FUNCTION_BLOCK Desinfeccao_UV (* Desinfeccao UV e limitacao da vazao de lancamento (700) - HidrycoLib *)
  (* Standard: 61499-2 *)
  (* Version 1.3, 21/10/2026, Hidryco, Hidryco, 1.3: REQ_GERADOR (geradorHabilitaUV01/02, stsGerador; Subestacao HAB_UV_700_01/02 e stsPlantaNoGerador) repassado ao UV para o raio dos canais. 1.2: pidCtl Pid com CycleTime 1000 ms (sem ele o calculo ciclico do pidSC ficava sem periodo). 1.1: ajustes do PID no sub-CAT PID_VC_700_01 (padrao Desinfeccao do legado; desejado = vazao maxima); reset cmdResetFalhas / E_RESET_FALHAS_PROCESSO; AIT_700_01/03/04. 1.0: desinfeccao (700). Sub-CATs: VC_700_01 (Valvula_Coester modulante), UV (UV_Trojan), FT_700_01 (Parshall 4-20 mA, m3/h), AIT_700_001 turbidez, AIT_700_003 pH, AIT_700_004 OD (SC4500 por comunicacao). PID continuo (pidCtl, Direction TRUE: vazao acima do setpoint fecha a valvula) limita a vazao de lancamento (padrao 1242 m3/h = 345 L/s). Campo por symlink ${PATH}: djPCEDesligado, djPCMDesligado, djUV01, djUV02, djVC01, djMO01 (remota %I0.0-0.5), stsRemotaComOk (COM_OK do IO_DI32 da remota). *)
  PACKAGE Hidryco.HidrycoLib;
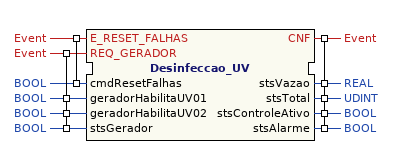
  EVENT_INPUT
    E_RESET_FALHAS WITH cmdResetFalhas; (* Reset pelo processo (desinfeccao, valvula, UV e sensores) com cmdResetFalhas = TRUE *)
    REQ_GERADOR WITH geradorHabilitaUV01, geradorHabilitaUV02, stsGerador; (* Planta no gerador e liberacao do UV (Subestacao) *)
  END_EVENT
  EVENT_OUTPUT
    CNF WITH stsVazao, stsTotal, stsControleAtivo, stsAlarme; (* Status *)
  END_EVENT
  VAR_INPUT
    cmdResetFalhas : BOOL; (* TRUE = reset (com o evento E_RESET_FALHAS) *)
    geradorHabilitaUV01 : BOOL; (* 700-UV-01 liberado para operar com a planta nos geradores *)
    geradorHabilitaUV02 : BOOL; (* 700-UV-02 liberado para operar com a planta nos geradores *)
    stsGerador : BOOL; (* TRUE = planta alimentada pelos geradores *)
  END_VAR
  VAR_OUTPUT
    stsVazao : REAL; (* Vazao do efluente final (m3/h) *)
    stsTotal : UDINT; (* Volume totalizado (m3) *)
    stsControleAtivo : BOOL; (* PID controlando a 700-VC-01 *)
    stsAlarme : BOOL; (* Algum alarme da desinfeccao *)
  END_VAR
  FBS
    IThis : Desinfeccao_UV_HMI(QI := TRUE);
    plcStart1 : plcStart(Prio := 10);
    Logica : basicDesinfeccao;
    Tick : E_CYCLE(DT := T#1s);
    Pid : pidCtl(CycleTime := 1000, Direction := TRUE, Bump := FALSE, ProhibitOutInc := FALSE, ProhibitOutDec := FALSE);
    PersTotal : PERSISTENCE_20652AC5DB8BA8AD5(QI := TRUE); {SET_ATTRIBUTE(Configuration.GenericFBType.InterfaceParams, Runtime.Standard#I:=3;input${I$}:UINT,UINT,UDINT)}
    Disjuntores : SYMLINKMULTIVARDST_5495E501E675F500(QI := TRUE, NAME1 := '$${PATH}djPCEDesligado', NAME2 := '$${PATH}djPCMDesligado', NAME3 := '$${PATH}djUV01', NAME4 := '$${PATH}djUV02', NAME5 := '$${PATH}djVC01', NAME6 := '$${PATH}djMO01'); {SET_ATTRIBUTE(Configuration.GenericFBType.InterfaceParams, Runtime.System#I:=6;VALUE${I$}:BOOL,BOOL,BOOL,BOOL,BOOL,BOOL)}
    Remota : SYMLINKMULTIVARDST_1559B0FF8170C9BA0(QI := TRUE, NAME1 := '$${PATH}stsRemotaComOk'); {SET_ATTRIBUTE(Configuration.GenericFBType.InterfaceParams, Runtime.System#I:=1;VALUE${I$}:BOOL)}
    FT_700_01 : Sensor_Generico(pin_CC8EEC06FF0C4430 := 'm3/h', pin_6D3A2524C5D0F0D1 := 0);
    AIT_700_01 : Sensor_Generico(pin_D46B37D45FD5AF5D := TRUE, pin_0ECE7B3867B02E0B := TRUE, pin_CC8EEC06FF0C4430 := 'NTU', pin_6D3A2524C5D0F0D1 := 1);
    AIT_700_03 : Sensor_Generico(pin_D46B37D45FD5AF5D := TRUE, pin_0ECE7B3867B02E0B := TRUE, pin_CC8EEC06FF0C4430 := '', pin_6D3A2524C5D0F0D1 := 2);
    AIT_700_04 : Sensor_Generico(pin_D46B37D45FD5AF5D := TRUE, pin_CC8EEC06FF0C4430 := 'mV', pin_6D3A2524C5D0F0D1 := 0); (* ORP (mV) do SC4500 de pH (conexao supervisionada pelo AIT_700_03: o connStatusInt so tem um destino) *)
    VC_700_01 : Atuador_Coester(pin_C65F121E4D57852C := TRUE);
    UV : UV_Trojan;
    AlarmeVazaoAlta : ALARM_BIT(TYPE := 1, ACKTYPE_1 := 2, ACTIVE := TRUE); {SET_ATTRIBUTE(HMI.AlarmText, Vazão de lançamento acima do limite)}
    AlarmeVariacao : ALARM_BIT(TYPE := 1, ACKTYPE_1 := 2, ACTIVE := TRUE); {SET_ATTRIBUTE(HMI.AlarmText, Variação brusca da vazão de lançamento)} {SET_ATTRIBUTE(HMI.AlarmClass, Warning)}
    AlarmeDisjuntor : ALARM_BIT(TYPE := 1, ACKTYPE_1 := 2, ACTIVE := TRUE); {SET_ATTRIBUTE(HMI.AlarmText, Disjuntor da desinfecção desligado)} {SET_ATTRIBUTE(HMI.AlarmClass, Warning)}
    AlarmeRemota : ALARM_BIT(TYPE := 1, ACKTYPE_1 := 2, ACTIVE := TRUE); {SET_ATTRIBUTE(HMI.AlarmText, Remota da desinfecção sem comunicação)} {SET_ATTRIBUTE(HMI.AlarmClass, Warning)}
    PID_VC_700_01 : Controle_PID;
  END_FBS
  EVENT_CONNECTIONS
    plcStart1.FIRST_INIT TO IThis.B18F9527B03F6368;
    plcStart1.REDO_INIT TO IThis.B18F9527B03F6368;
    IThis.8DA18C8B88D861AA TO Disjuntores.INIT;
    Disjuntores.INITO TO Remota.INIT;
    Remota.INITO TO Logica.9E12B42E11EB9FB7;
    Remota.INITO TO IThis.B29E261CF0325DC9;
    Logica.39B67DFC9697D1D0 TO Tick.START;
    Logica.39B67DFC9697D1D0 TO PersTotal.INIT;
    PersTotal.INITO TO PersTotal.READ;
    PersTotal.READCNF TO Logica.2E96492E37281113;
    Logica.BC4C937414AD6E45 TO PersTotal.WRITE;
    Logica.39B67DFC9697D1D0 TO AlarmeVazaoAlta.INIT;
    AlarmeVazaoAlta.INITO TO AlarmeVazaoAlta.REQ_INITDATA;
    AlarmeVazaoAlta.CNF_INITDATA TO AlarmeVazaoAlta.ACTIVATE;
    AlarmeVariacao.INITO TO AlarmeVariacao.REQ_INITDATA;
    AlarmeVariacao.CNF_INITDATA TO AlarmeVariacao.ACTIVATE;
    AlarmeVazaoAlta.INITO TO AlarmeVariacao.INIT;
    AlarmeDisjuntor.INITO TO AlarmeDisjuntor.REQ_INITDATA;
    AlarmeDisjuntor.CNF_INITDATA TO AlarmeDisjuntor.ACTIVATE;
    AlarmeVariacao.INITO TO AlarmeDisjuntor.INIT;
    AlarmeRemota.INITO TO AlarmeRemota.REQ_INITDATA;
    AlarmeRemota.CNF_INITDATA TO AlarmeRemota.ACTIVATE;
    AlarmeDisjuntor.INITO TO AlarmeRemota.INIT;
    AlarmeRemota.INITO TO plcStart1.ACK_FIRST;
    Tick.EO TO Logica.A43A58424E0F5DF5;
    Disjuntores.CNF TO Logica.22B807AE7A8B903D;
    Remota.CNF TO Logica.2AE8EBA1815E0012;
    FT_700_01.28A380156DB271B8 TO Logica.6559A273E8431D42;
    VC_700_01.CF6616D3CB5312F6 TO Logica.4F5B69463931E86B;
    UV.41148E14CCAE49D5 TO Logica.1495D2B4E524DEC3;
    Logica.6010724B5A00E1A3 TO VC_700_01.6AE7937B5439A162;
    FT_700_01.28A380156DB271B8 TO Pid.REQ;
    Logica.38355A458523F08C TO Pid.REQ;
    Pid.CNF TO Logica.1DD56BE62400BF1C;
    Pid.C_CNF TO Logica.1DD56BE62400BF1C;
    IThis.341E4C9D143B2914 TO Logica.69B239DBC6B5BF03;
    IThis.673C9CACFA30E81B TO Logica.F980CDC9B2AFA9D8;
    IThis.A7123D0B6BA18805 TO Logica.B454118112B7B3A8;
    Logica.04CB25776C0D242A TO IThis.1B47BC94CEE432D9;
    Logica.04CB25776C0D242A TO AlarmeVazaoAlta.REQ;
    AlarmeVazaoAlta.IND_1 TO IThis.1B47BC94CEE432D9;
    IThis.673C9CACFA30E81B TO AlarmeVazaoAlta.ACK_C1;
    Logica.04CB25776C0D242A TO AlarmeVariacao.REQ;
    AlarmeVariacao.IND_1 TO IThis.1B47BC94CEE432D9;
    IThis.673C9CACFA30E81B TO AlarmeVariacao.ACK_C1;
    Logica.04CB25776C0D242A TO AlarmeDisjuntor.REQ;
    AlarmeDisjuntor.IND_1 TO IThis.1B47BC94CEE432D9;
    IThis.673C9CACFA30E81B TO AlarmeDisjuntor.ACK_C1;
    Logica.04CB25776C0D242A TO AlarmeRemota.REQ;
    AlarmeRemota.IND_1 TO IThis.1B47BC94CEE432D9;
    IThis.673C9CACFA30E81B TO AlarmeRemota.ACK_C1;
    E_RESET_FALHAS TO Logica.DA13244B5D56E79F;
    E_RESET_FALHAS TO FT_700_01.D21DAA5004F58516;
    E_RESET_FALHAS TO AIT_700_01.D21DAA5004F58516;
    E_RESET_FALHAS TO AIT_700_03.D21DAA5004F58516;
    E_RESET_FALHAS TO AIT_700_04.D21DAA5004F58516;
    E_RESET_FALHAS TO VC_700_01.D903CD18EBE204D1;
    Logica.6AA932C3761CE99C TO CNF;
    PID_VC_700_01.75EB05A15DC6DC61 TO Pid.REQ_PARA;
    PID_VC_700_01.75EB05A15DC6DC61 TO Pid.REQ_SP;
    PID_VC_700_01.75EB05A15DC6DC61 TO Logica.69B239DBC6B5BF03;
    Remota.INITO TO PID_VC_700_01.117942CC3F34C94C;
    Logica.04CB25776C0D242A TO PID_VC_700_01.7BD84B0FC1882775;
    REQ_GERADOR TO UV.6FAFCDDE653CB65D;
  END_CONNECTIONS
  DATA_CONNECTIONS
    PersTotal.output3 TO Logica.E77A551E7F1625D6;
    Logica.BB35FC69145014F5 TO PersTotal.input3;
    Disjuntores.VALUE1 TO Logica.CF45361D95BFAA25;
    Disjuntores.VALUE2 TO Logica.347EEF72575B0DAD;
    Disjuntores.VALUE3 TO Logica.159FAE7A20FE4F43;
    Disjuntores.VALUE4 TO Logica.7868F97BB44D7BB6;
    Disjuntores.VALUE5 TO Logica.92824DDB3BCC4699;
    Disjuntores.VALUE6 TO Logica.50FED92E4734ACF3;
    Remota.VALUE1 TO Logica.D0484A6EFE322016;
    FT_700_01.D7422D307E6AF52D TO Logica.F569AB39D886D3C5;
    FT_700_01.726640D1704B3F86 TO Logica.8F6D70C85B5729EE;
    VC_700_01.904DD3246D8E0F2F TO Logica.C5936F826382DFB8;
    VC_700_01.259F220E31BE1DFA TO Logica.7315FEF776808725;
    VC_700_01.5B46E3B5D12031DA TO Logica.023A1B52E4E2056D;
    VC_700_01.378CDAA06C4824E3 TO Logica.DBD5C62FC984909D;
    UV.8A986F32247F8461 TO Logica.DB1DCC8BAF4C9029;
    UV.EDFBC67855FC1BF4 TO Logica.1AFFBF765DAF6E05;
    UV.53F24ADA26C29448 TO Logica.6927441A48A28A44;
    UV.E73DB33437F0D160 TO Logica.FA4C9F16C9AD1E00;
    UV.B5E6F2B1B4A7F74D TO Logica.E17D46372D8AC1CC;
    UV.2373201554B21091 TO Logica.CA02F082C523342B;
    Logica.635B91EC32B193D8 TO VC_700_01.B08C4ED4004BD1E2;
    FT_700_01.D7422D307E6AF52D TO Pid.Pv;
    Logica.B925699CCA1010B0 TO Pid.Mode;
    Logica.E0C52E4AA1CB94A3 TO Pid.PresetValue;
    Pid.Out TO Logica.AA3C6B9770CFA1D6;
    IThis.975D7F4B71294A99 TO Logica.A62BE056EBF6633F;
    IThis.48B1DA7F68ECA0A8 TO Logica.0CA93D1DC0F0D80A;
    IThis.BF0DC1C37334FADC TO Logica.EAB397A6710197DE;
    IThis.3223A03025B9D306 TO Logica.14F8441489A49AD8;
    IThis.133D4C207A85139E TO Logica.EDA9F4A4D8516735;
    Logica.8B489663C97AF746 TO IThis.64C5B4D669700647;
    Logica.2CB6FFAA3F88FD37 TO IThis.9BBBF4F79C014F9D;
    Logica.1AC4273BD48629B4 TO IThis.ED2A3A2AD9D2CEAB;
    Logica.7C47B967196CD681 TO IThis.8CFA6BB1EE69DBDA;
    Logica.F5E44B9CD467E225 TO IThis.9D544CFE60C51E40;
    Logica.E0E853656DE9663A TO IThis.00083F484189930B;
    Logica.5B994E1E72A57859 TO IThis.5A630CE8F223E31A;
    Logica.9D46B9FE82DC9AB1 TO IThis.3724F9189B78EC4D;
    Logica.06E435E0579C0A31 TO IThis.4C496D880FB42A44;
    Logica.03E13841379C7979 TO IThis.DE11125D4105DF0E;
    Logica.9EE277DF1A6EE639 TO IThis.909A978770157DD8;
    Logica.DD39785BA0B3D6D1 TO IThis.D8676A9461C485D9;
    Logica.DC6A854DD28F4447 TO IThis.8155290424886535;
    Logica.CFF2FF9B070BCB84 TO IThis.E0FD426C54E10B50;
    Logica.A1948102A71BA04F TO IThis.B5278628A6F4EB0E;
    Logica.49CC92A2C50C5502 TO IThis.3146A9607323897C;
    Logica.029A5972D76D7D9D TO IThis.207239DB8C69408E;
    Logica.7C31ABB79E620CA1 TO IThis.0DCEC12DB41BD8A9;
    Logica.4979C9EBFE656646 TO IThis.F89132E9AC0FBE71;
    Logica.9AA3D7C962B2722B TO IThis.A35FB648721D6941;
    Logica.F5BC914DFDB76B1B TO IThis.2B50411206C948D5;
    Logica.2E78B7E52A0ED234 TO IThis.8B80C37723B8B9A9;
    Logica.C779F990E9DA2177 TO IThis.946F4BE0E36C2836;
    Logica.9AA3D7C962B2722B TO AlarmeVazaoAlta.INP;
    AlarmeVazaoAlta.STATE_1 TO IThis.060041ABB2A0A5A2;
    Logica.F5BC914DFDB76B1B TO AlarmeVariacao.INP;
    AlarmeVariacao.STATE_1 TO IThis.3988E692C5278158;
    Logica.4979C9EBFE656646 TO AlarmeDisjuntor.INP;
    AlarmeDisjuntor.STATE_1 TO IThis.F7176D1924986299;
    Logica.2E78B7E52A0ED234 TO AlarmeRemota.INP;
    AlarmeRemota.STATE_1 TO IThis.6D5DB80D1692E5C6;
    cmdResetFalhas TO Logica.5A0059668713CC5A;
    cmdResetFalhas TO FT_700_01.1908F43CB878F5E7;
    cmdResetFalhas TO AIT_700_01.1908F43CB878F5E7;
    cmdResetFalhas TO AIT_700_03.1908F43CB878F5E7;
    cmdResetFalhas TO AIT_700_04.1908F43CB878F5E7;
    cmdResetFalhas TO VC_700_01.C82CBBE25FC56079;
    Logica.8B489663C97AF746 TO stsVazao;
    Logica.2C19FD8E73A079CA TO stsTotal;
    Logica.7C47B967196CD681 TO stsControleAtivo;
    Logica.C779F990E9DA2177 TO stsAlarme;
    PID_VC_700_01.C9DF845DD1ECA932 TO Pid.Sp;
    PID_VC_700_01.C9DF845DD1ECA932 TO Logica.3EF61F60D9980F84;
    PID_VC_700_01.4F45CBCE24FA8775 TO Pid.Gain;
    PID_VC_700_01.5D86C7647B367BF7 TO Pid.IntegralTime;
    PID_VC_700_01.C753842CF6C65D61 TO Pid.DerivativeTime;
    PID_VC_700_01.8B11A5B11AA557C3 TO Pid.OutMin;
    PID_VC_700_01.8B11A5B11AA557C3 TO Logica.DF73D60158F656E4;
    PID_VC_700_01.E7AF90225A9267BD TO Pid.OutMax;
    PID_VC_700_01.E7AF90225A9267BD TO Logica.0F4CFB3D37BB8386;
    PID_VC_700_01.004F03C1536C2B1E TO Logica.FEC6CBE54CA37A44;
    Logica.BB5C6CDA218388F6 TO PID_VC_700_01.260D6E81A1639D84;
    geradorHabilitaUV01 TO UV.29A04DF02BFCF18C;
    geradorHabilitaUV02 TO UV.410574851060558C;
    stsGerador TO UV.9B4A40E24325447A;
  END_CONNECTIONS
END_FUNCTION_BLOCK
